Staubli VAL3: robotStatus.pjx

--- robotStatus.pjx ---
Parameters version=s8.21cs9_BS4703 stackSize=200000 millimeterUnit=true
Program file=addLog.pgx
Program file=getAlarmMsg.pgx
Program file=getLog.pgx
Program file=init.pgx
Program file=resetAlarm.pgx
Program file=robotStatus.pgx
Program file=saveLog.pgx
Program file=setAlarm.pgx
Program file=start.pgx
Program file=stop.pgx
Data file=robotStatus.dtx
Library alias=Log path=./log/log.pjx autoload=true password=

--- robotStatus.dtx ---
public bool _bHeavyAlarm
public bool bAlarmAck
public bool bGOTO
public bool bInSwitch
public bool bIsCycle
public bool bIsError
public bool bIsEstop
public bool bIsHome
public bool bIsMoving
public bool bIsPause
public bool bIsReady
public bool bIsRemoteAuto
public bool bIsSaving
public bool bPowerON
public bool bProgGOTO
public bool bQuitApp
public bool bReloadIO
public bool bSimulate
public bool bToPause
public bool bToStartCycle
public bool bToStopCycle
public num _nAlarmCode[10] = 300
num _nAlarmIndex
public num _nAvgCapacity
public num _nBestCapacity
public num _nCTIndex
public num _nCapacity
public num _nCycleTime
public num _nErrIndex[10]
  [1] = -1
  [2] = -1
  [3] = -1
  [4] = -1
  [5] = -1
  [6] = -1
  [7] = -1
  [8] = -1
  [9] = -1
public num _nOmacStat = 9
public num nActCode
public num nCycleCmd
public num nCycleIndex = 78
public num nCycleMoveID
public num nFrameIndex
public num nHMIcmd
public num nHWState
public num nHeavyAlarmLev
public num nPLCcmd
public num nProgCode = 4
public num nProgFb = 1
public num nSetSwitchValue
public num nToolIndex
public num nTrajCode
public string _sRobotStatus = "错误：-300. :0traj数据库加载错误"
public string sAlarmMes[10]
public string sBusUsing = "PROFINET"
public string sCycleItem = "04 sls"
public string sIOStatus
string sLstIOStatus
string sLstRobStatus
string sLstTrajStatus
public string sPageUsing
public string sTrajStatus = "[04 sls]移动到:78, DOUT[11]-喷涂完成=FALSE"

--- start.pgx ---
program start()
begin
end

--- _clickIoPage.pgx ---
public program _clickIoPage()
begin
  sPageUsing="InOut"
  userPage("Disk://source/projectSource/io/interface/InOut")
  delay(1)
end

--- _clickProductionPage.pgx ---
public program _clickProductionPage()
begin
  sPageUsing="cycleCtrl"
  userPage("Disk://Project/interface/cycleCtrl")
  delay(1)
end

--- addLog.pgx ---
public program addLog(string x_sLog (dimensions=1), num x_nType (dimensions=1))
begin
  call Log:addlog(x_sLog,x_nType)
end

--- getAlarmMsg.pgx ---
program getAlarmMsg(num x_nAlarmCode (dimensions=1), string& x_sMsg (dimensions=1))
begin
  //
  switch x_nAlarmCode
    //**************************************动作************************************
    case 200
      x_sMsg=".8"
    break
    case 201
      x_sMsg="动作堆栈溢出，无法执行最新动作"
    break
    case 202
      x_sMsg="动作百分比错误"
    break
    case 203
      x_sMsg="动作中的输入输出的InOutType类型错误"
    break
    case 204
      x_sMsg="动作中的输入输出的输入输出索引号错误"
    break
    case 205
      x_sMsg="动作中的输入输出的输出值参数错误"
    break
    case 206
      x_sMsg="动作中的输入输出的脉冲时间参数值错误"
    break
    case 207
      x_sMsg="动作中的输入输出的输入值参数值错误"
    break
    case 208
      x_sMsg="动作的范围超限"
    break
    case 209
      x_sMsg="动作错误"
    break
    case 210
      x_sMsg=".8"
    break


    //*************************************点位超限**************************************
    case 220
      x_sMsg="Point点位超限"
    break
    case 221
      x_sMsg="Joint点位超限"
    break
    case 300
      x_sMsg="traj数据库加载错误"
    break
    case 301
      x_sMsg="prog数据库加载错误"
    break
    case 302
      x_sMsg="索引指向的数据库不存在"
    break
    case 303
      x_sMsg="自动运行过程中伺服异常下电"
    break
    ////*************************************系统报错**************************************
    case 400
      x_sMsg="[硬件报错]-电源错误,错误代码:"+toString(".8",nHWState)
    break
    case 401
      x_sMsg="[硬件报错]-RSI9错误,错误代码:"+toString(".8",nHWState)
    break
    case 402
      x_sMsg="[硬件报错]-STARC/DSI错误,错误代码:"+toString(".8",nHWState)
    break
    case 403
      x_sMsg="[硬件报错]-编码器错误,错误代码:"+toString(".8",nHWState)
    break
    case 404
      x_sMsg="[硬件报错]-驱动器错误,错误代码:"+toString(".8",nHWState)
    break
    case 405
      x_sMsg="[硬件报错]-手柄未安装,错误代码:"+toString(".8",nHWState)
    break
  endSwitch

end

--- getLog.pgx ---
public program getLog(string& x_sLog[] (dimensions=1), num x_nType (dimensions=1))
begin
  call Log:getlog(x_sLog,x_nType)
end

--- init.pgx ---
public program init()
begin
  //init all
  bIsSaving=false
  call resetAlarm()
  bAlarmAck=false
  bGOTO=false
  bIsCycle=false
  bIsEstop=false
  bIsHome=false
  bIsReady=false
  bReloadIO=false
  bSimulate=false
  bSimulate=false
  _bHeavyAlarm=false
  bQuitApp=false
  nCycleCmd=0
  nCycleMoveID=0
  nFrameIndex=0
  nHeavyAlarmLev=0
  nHMIcmd=0
  nPLCcmd=0
  nToolIndex=0
  _nAlarmIndex=0
  _nAvgCapacity=0
  _nBestCapacity=0
  _nCapacity=0
  _nCTIndex=0
  _nCycleTime=0
  _nOmacStat=9

  sPageUsing=""
  sTrajStatus=""
  sLstTrajStatus=""
  _sRobotStatus=""
  sLstRobStatus=""
  sIOStatus=""
  sLstIOStatus=""

end

--- resetAlarm.pgx ---
public program resetAlarm()
  local num l_n
begin
  for l_n=0 to size(_nAlarmCode)-1
    _nErrIndex[l_n]=-1
    _nAlarmCode[l_n]=0
    sAlarmMes[l_n]=""
  endFor
  _nAlarmIndex=0
end

--- robotStatus.pgx ---
public program robotStatus()
begin
  //检测状态显示变化
  if _sRobotStatus!=sLstRobStatus
    sLstRobStatus=_sRobotStatus
    call Log:addlog(toString(".3",clock())+" "+"[状态信息]:"+_sRobotStatus+getDate(" %m-%d %H:%M:%S"),1)
  endIf

  if sTrajStatus!=sLstTrajStatus
    sLstTrajStatus=sTrajStatus
    call Log:addlog(toString(".3",clock())+" "+"[路径信息]:"+sTrajStatus+getDate(" %m-%d %H:%M:%S"),2)
  endIf

  if sIOStatus!=sLstIOStatus
    sLstIOStatus=sIOStatus
    call Log:addlog(toString(".3",clock())+" "+"[信号信息]:"+sIOStatus+getDate(" %m-%d %H:%M:%S"),3)
  endIf
end

--- saveLog.pgx ---
public program saveLog(string x_sPath (dimensions=1), num& x_nResult (dimensions=1))
  local num l_n
  local num l_nLogMsgIndex
begin
  if x_sPath==""
    x_nResult=Log:libSave()
  else
    x_nResult=Log:libSave(x_sPath)
  endIf
  delay(0.5)
end

--- setAlarm.pgx ---
public program setAlarm(num x_nAlarmCode (dimensions=1), num x_nErrIndex (dimensions=1))
  local bool l_bExist
  local num l_nIndex
  local string l_sAlarmLevel
  local string l_sErrMsg
begin
  //check if the alarm has existed in the list
  do
    l_bExist=(x_nAlarmCode==_nAlarmCode[l_nIndex] and x_nErrIndex==_nErrIndex[l_nIndex])
    l_nIndex=l_nIndex+1
  until l_bExist or l_nIndex>=size(_nAlarmCode)
  //
  if !l_bExist
    //new alarm, add it
    if _nAlarmCode[_nAlarmIndex]>0
      _nAlarmIndex=(_nAlarmIndex+1)%size(_nAlarmCode)
    endIf
    _nAlarmCode[_nAlarmIndex]=x_nAlarmCode
    _nErrIndex[_nAlarmIndex]=x_nErrIndex
    call getAlarmMsg(x_nAlarmCode,l_sErrMsg)
    //错误等级
    if _nAlarmCode[_nAlarmIndex]>=0
      if x_nAlarmCode>nHeavyAlarmLev
        l_sAlarmLevel="错误："
      else
        l_sAlarmLevel="警告："
      endIf
      //错误消息
      if x_nErrIndex>=0
        sAlarmMes[_nAlarmIndex]=_sRobotStatus=l_sAlarmLevel+"-"+toString("",x_nAlarmCode)+". "+":"+toString("",x_nErrIndex)+l_sErrMsg
      else
        sAlarmMes[_nAlarmIndex]=_sRobotStatus=l_sAlarmLevel+"-"+toString("",x_nAlarmCode)+". "+l_sErrMsg
      endIf
      logMsg(sAlarmMes[_nAlarmIndex])
    endIf
    delay(0)
  endIf
end

--- stop.pgx ---
program stop()
begin
end
